{region 'Documentation'}
(*!
<summary>Checks that at least one selected bit is TRUE.</summary>
*)
{endregion}
FUNCTION_BLOCK AssertContainsTrue_Byte EXTENDS AssertionBase
VAR_INPUT
    IN : BYTE; //! Actual bitfield.
    Mask : BYTE := 16#FF; //! Selects evaluated bits; defaults to all bits. An empty mask produces Error during evaluation.
END_VAR

SUPER^();

{region 'Documentation'}
(*!
<summary>Rejects an empty mask before checking for a matching selected bit.</summary>
*)
{endregion}
METHOD PROTECTED Assert
VAR
    Message : STRING(GVL_Constants.MessageLength);
    MaskText : STRING(GVL_Constants.AssertionValueLength);
    ActualText : STRING(GVL_Constants.AssertionValueLength);
END_VAR
VAR CONSTANT
    NoMask : BYTE := 16#00;
    HexDigitCount : USINT := 2;
END_VAR
IF NOT EvaluationActive THEN
    RETURN;
END_IF;

IF Result = E_Result.Error THEN
    RETURN;
END_IF;

IF Mask = NoMask THEN
    MaskText := CreateAssertionTextValue_Hex(Value := BYTE_TO_LWORD(Mask),
        DigitCount := HexDigitCount);
    Message := CONCAT('Assertion error: mask must not be empty. Mask = ',
        MaskText);
    Message := CONCAT(Message, '.');
    Error(Message := Message);
    RETURN;
END_IF;

IF Result = E_Result.Failed THEN
    RETURN;
END_IF;

IF (IN AND Mask) = NoMask THEN
    MaskText := CreateAssertionTextValue_Hex(Value := BYTE_TO_LWORD(Mask),
        DigitCount := HexDigitCount);
    ActualText := CreateAssertionTextValue_Hex(Value := BYTE_TO_LWORD(IN),
        DigitCount := HexDigitCount);
    Message := CONCAT('Assertion failed: no selected bit is TRUE. Mask = ',
        MaskText);
    Message := CONCAT(Message, ', Actual = ');
    Message := CONCAT(Message, ActualText);
    Message := CONCAT(Message, '.');
    Fail(Message := Message);
    RETURN;
END_IF;

Pass();
END_METHOD

END_FUNCTION_BLOCK

(* stored: Version 1.1.0.1
   POU AssertContainsTrue_Byte: Id {9db78fd3-9e56-4668-8995-bd3e6bb59b3d}, SpecialFunc None
   Folder Internal: Id {49c1e5ad-9b06-4965-8f23-62d2314e09e3}
   Method Assert: Id {78eac5bd-19f5-499f-a430-e9f7528dd118} *)
